ADAPTER buttons_manual (* Adapter Interface *)
  (* Standard: 61499-1 *)
  (* Version 0.0, 10/22/2026, macie, Schneider Electric *)
  PACKAGE Main;
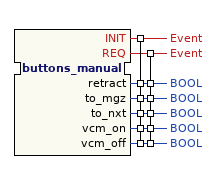
  EVENT_OUTPUT
    INIT WITH retract, to_mgz, to_nxt, vcm_on, vcm_off;
    REQ WITH retract, to_mgz, to_nxt, vcm_on, vcm_off;
  END_EVENT
  VAR_OUTPUT
    retract : BOOL;
    to_mgz : BOOL;
    to_nxt : BOOL;
    vcm_on : BOOL;
    vcm_off : BOOL;
  END_VAR
  SERVICE SOCKET/PLUG
    SEQUENCE request_confirm
      SOCKET.REQ(retract) -> PLUG.REQ(retract);
      PLUG.CNF(CNFD) -> SOCKET.CNF(CNFD);
    END_SEQUENCE
    SEQUENCE indication_response
      PLUG.IND(INDD) -> SOCKET.IND(INDD);
      SOCKET.RSP(to_mgz) -> PLUG.RSP(to_mgz);
    END_SEQUENCE
  END_SERVICE
END_ADAPTER
